(* IEC 61131-3 sources: RootPLC/conformance/cases/test-blocks, 12 files *)

(* ---- ok_asserts.st ---- *)
(* spec: [tests.assert] [pous.test]
   expect: ok *)
FUNCTION Add : INT
VAR_INPUT
    a, b : INT;
END_VAR
Add := a + b;
END_FUNCTION

TEST add_works
VAR
    r : INT;
END_VAR
r := Add(2, 3);
ASSERT_EQ(5, r);
ASSERT_NE(4, r);
ASSERT_TRUE(r > 0);
ASSERT_FALSE(r < 0);
END_TEST

(* ---- err_private_outside_test.st ---- *)
(* spec: [tests.whitebox] [pous.call.local-read]
   expect: error RP0203 *)
FUNCTION_BLOCK FB_Count
VAR
    hidden : INT;
END_VAR
END_FUNCTION_BLOCK

PROGRAM PRG_Main
VAR
    c : FB_Count;
    n : INT;
END_VAR
c.hidden := n;   (* outside a TEST block internal variables are read-only *)
END_PROGRAM

(* ---- ok_evidence_no_tests.st ---- *)
(* spec: [tests.evidence]
   expect: ok
   evidence: not verified *)
(* A program without TEST blocks compiles, but nothing has been verified. *)
FUNCTION_BLOCK FB_Latch
VAR_INPUT
    start : BOOL;
    stop : BOOL;
END_VAR
VAR_OUTPUT
    running : BOOL;
END_VAR
running := (start OR running) AND NOT stop;
END_FUNCTION_BLOCK

(* ---- ok_evidence_verified.st ---- *)
(* spec: [tests.evidence] [tests.mutation]
   expect: ok
   mutate: killed=3 viable=3
   evidence: verified *)
FUNCTION_BLOCK FB_Latch
VAR_INPUT
    start : BOOL;
    stop : BOOL;
END_VAR
VAR_OUTPUT
    running : BOOL;
END_VAR
running := (start OR running) AND NOT stop;
END_FUNCTION_BLOCK

TEST latch_sets_holds_and_stops
VAR
    l : FB_Latch;
END_VAR
l(start := TRUE, stop := FALSE);
ASSERT_TRUE(l.running);
l(start := FALSE, stop := FALSE);
ASSERT_TRUE(l.running);
l(start := TRUE, stop := TRUE);
ASSERT_FALSE(l.running);
END_TEST

(* ---- ok_mutation_all_killed.st ---- *)
(* spec: [tests.mutation]
   expect: ok
   mutate: killed=3 viable=3 *)
FUNCTION_BLOCK FB_Latch
VAR_INPUT
    start : BOOL := FALSE;
    stop : BOOL := FALSE;
END_VAR
VAR_OUTPUT
    running : BOOL;
END_VAR
running := (start OR running) AND NOT stop;
END_FUNCTION_BLOCK

TEST latch_sets_holds_and_stops
VAR
    l : FB_Latch;
END_VAR
l(start := TRUE, stop := FALSE);
ASSERT_TRUE(l.running);
l(start := FALSE, stop := FALSE);
ASSERT_TRUE(l.running);
l(start := TRUE, stop := TRUE);
ASSERT_FALSE(l.running);
END_TEST

(* ---- ok_mutation_operators.st ---- *)
(* spec: [tests.mutation]
   expect: ok
   mutate: killed=5 viable=5 *)
FUNCTION_BLOCK FB_Level
VAR_INPUT
    level : INT;
END_VAR
VAR_OUTPUT
    high : BOOL;
    margin : INT;
    alarm : BOOL;
END_VAR
VAR
    t : TON;
END_VAR
high := level >= 80;
margin := 100 - level;
t(IN := high, PT := T#2s);
alarm := t.Q;
END_FUNCTION_BLOCK

TEST level_limits
VAR
    f : FB_Level;
END_VAR
f(level := 79);
ASSERT_FALSE(f.high);
ASSERT_EQ(21, f.margin);
f(level := 80);
ASSERT_TRUE(f.high);
ASSERT_EQ(20, f.margin);
ADVANCE(T#2s);
f(level := 80);
ASSERT_TRUE(f.alarm);
END_TEST

TEST alarm_not_early
VAR
    f : FB_Level;
END_VAR
f(level := 90);
ADVANCE(T#3s);
f(level := 90);
ASSERT_TRUE(f.alarm);
ADVANCE(T#1s);
END_TEST

(* ---- ok_mutation_survivor.st ---- *)
(* spec: [tests.mutation]
   expect: ok
   mutate: killed=2 viable=3 *)
FUNCTION_BLOCK FB_Latch
VAR_INPUT
    start : BOOL;
    stop : BOOL;
END_VAR
VAR_OUTPUT
    running : BOOL;
END_VAR
running := (start OR running) AND NOT stop;
END_FUNCTION_BLOCK

(* This test never checks stop, so replacing AND by OR survives. *)
TEST latch_sets
VAR
    l : FB_Latch;
END_VAR
l(start := TRUE, stop := FALSE);
ASSERT_TRUE(l.running);
END_TEST

(* ---- ok_tests_slice.st ---- *)
(* spec: [tests.slice]
   expect: ok *)
(* With rootplc test --slice, this file (it has a TEST block) and the files
   declaring what it uses are compiled; other files of the project are left
   out, also when they do not compile (crates/rootplc-driver/tests/
   test_slice.rs). *)
FUNCTION_BLOCK FB_Counter
VAR_INPUT up : BOOL; END_VAR
VAR_OUTPUT n : INT; END_VAR
VAR e : R_TRIG; END_VAR
e(CLK := up);
IF e.Q THEN
    n := n + 1;
END_IF;
END_FUNCTION_BLOCK

TEST counter_counts_edges
VAR c : FB_Counter; END_VAR
c(up := TRUE);
c(up := TRUE);
c(up := FALSE);
c(up := TRUE);
ASSERT_EQ(2, c.n);
END_TEST

(* ---- ok_whitebox.st ---- *)
(* spec: [tests.whitebox] [tests.runner]
   expect: ok *)
FUNCTION_BLOCK FB_Count
VAR_INPUT
    pulse : BOOL;
END_VAR
VAR
    hidden : INT;
END_VAR
IF pulse THEN
    hidden := hidden + 1;
END_IF;
END_FUNCTION_BLOCK

TEST internal_state_is_visible
VAR
    uut : FB_Count;
END_VAR
uut(pulse := TRUE);
uut(pulse := TRUE);
ASSERT_EQ(2, uut.hidden);
END_TEST

(* ---- err_advance_outside_test.st ---- *)
(* spec: [tests.time]
   expect: error RP0203 *)
PROGRAM PRG_Main
ADVANCE(T#1s);
END_PROGRAM

(* ---- err_assert_not_bool.st ---- *)
(* spec: [tests.assert]
   expect: error RP0103 *)
TEST bad_assert
VAR
    i : INT := 1;
END_VAR
ASSERT_TRUE(i);
END_TEST

(* ---- ok_advance_time.st ---- *)
(* spec: [tests.time]
   expect: ok *)
PROGRAM PRG_Alarm
VAR_INPUT
    high : BOOL;
END_VAR
VAR_OUTPUT
    alarm : BOOL;
END_VAR
VAR
    t : TON;
END_VAR
t(IN := high, PT := T#5s);
alarm := t.Q;
END_PROGRAM

TEST alarm_after_five_seconds
VAR
    uut : PRG_Alarm;
END_VAR
uut(high := TRUE);
ADVANCE(T#4s);
uut(high := TRUE);
ASSERT_FALSE(uut.alarm);
ADVANCE(T#1s);
uut(high := TRUE);
ASSERT_TRUE(uut.alarm);
ADVANCE(LT#1h);
uut(high := FALSE);
ASSERT_FALSE(uut.alarm);
END_TEST
